(* IEC 61131-3 sources: Test-Git_ESME26/TestProgettoESME_26.fbsproj/PacDriveLib Migration/Motion/MultiCam/PDL_FB_MultiCam.fb.st^/Init, 2 files *)

(* ---- Init.meth.st ---- *)
METHOD PRIVATE Init : BOOL
VAR_INPUT
END_VAR

Init := FALSE;

//check axis
IF i_ifDrive = 0 THEN
	SetDiagOutput(	i_etDiag	:= GD.ET_Diag.InputParameterInvalid,
					i_etDiagExt := PDL_ET_DiagExt.DriveInvalid,
					i_sMsg		:= 'i_ifDrive - Invalid Interface');
	RETURN;

ELSIF iq_lencMaster = 0 THEN
	SetDiagOutput(	i_etDiag	:= GD.ET_Diag.InputParameterInvalid,
					i_etDiagExt := PDL_ET_DiagExt.DriveInvalid,
					i_sMsg		:= 'iq_lencMaster - Invalid Interface');
	RETURN;
ELSE
	//get IF_DriveConfig
	xSuccess := __QUERYINTERFACE(i_ifDrive, ifGetParentDevice);
	IF xSuccess AND ifGetParentDevice <> 0 THEN
		ifDeviceAccess := ifGetParentDevice.GetParentDevice();
		xSuccess := __QUERYINTERFACE( ifDeviceAccess, ifDriveConfigAccess );
		IF xSuccess AND ifDriveConfigAccess <> 0 THEN
			ifDriveConfig := ifDriveConfigAccess.DriveConfig;
		END_IF
	END_IF

	xSuccess := __QUERYINTERFACE(ifDeviceAccess, ifDeviceTreeObjectAccess);
	IF xSuccess THEN
		sDriveName := ifDeviceTreeObjectAccess.DeviceTreeObject.Name;
	ELSE
		sDriveName := 'Axis';
	END_IF

	fbHalt.Axis := i_ifDrive;
	fbStop.Axis := i_ifDrive;
	fbMoveAbsolute.Axis := i_ifDrive;
	fbCamIn.Slave := i_ifDrive;
	fbCamIn.Master := iq_lencMaster;
	fbCamIn2.Slave := i_ifDrive;
	fbCamIn2.Master := iq_lencMaster;

	xSlaveIsModulo := i_ifDrive.xIsModulo;

END_IF

//read cycle time
pstTaskInfo := __CURRENTTASK.pTaskInfo;
IF pstTaskInfo <> 0
THEN
	lrOwnPlcTaskInterval	:= DWORD_TO_LREAL(pstTaskInfo^.dwInterval) / 1000000.0; //usec to sec
	lrTSwitch				:= DINT_TO_LREAL(i_diTXend) / 1000.0 + lrOwnPlcTaskInterval;
ELSE
	SetDiagOutput(	i_etDiag	:= GD.ET_Diag.UnexpectedProgramBehavior,
					i_etDiagExt := PDL_ET_DiagExt.UnexpectedFeedback,
					i_sMsg		:= 'IecTaskGetInfo3 - reading cycle time failed');
	RETURN;
END_IF

Init := TRUE;

(* ---- RegisterLoggerPoint.meth.st ---- *)
METHOD PUBLIC RegisterLoggerPoint
VAR_INPUT
	i_ifParent		: APL.IF_LoggerPoint;
	i_sName			: STRING[80];
END_VAR
VAR_OUTPUT
	q_etDiag		: GD.ET_Diag := GD.ET_Diag.Ok;
	q_etDiagExt		: PDL_ET_DiagExt := PDL_ET_DiagExt.Ok;
END_VAR
VAR
	etDiagBuffer		: GD.ET_Diag;
	etDiagExtBufferAPL	: APL.ET_DiagExt;
END_VAR

THIS^.fbLoggerPoint.RegisterLoggerPoint(	i_ifParent		:= i_ifParent,
											i_sName			:= i_sName,
											i_sType			:= 'FB_MultiCam',
											i_sSource		:= 'PDL',
											q_etDiag		=> etDiagBuffer,
											q_etDiagExt		=> etDiagExtBufferAPL);

IF (etDiagBuffer <> GD.ET_Diag.Ok) THEN
	CASE etDiagExtBufferAPL OF
		APL.ET_DiagExt.ParentInvalid:
			q_etDiag := GD.ET_Diag.InputParameterInvalid;
			q_etDiagExt := PDL_ET_DiagExt.ParentInvalid;

		APL.ET_DiagExt.ParentNotRegistered:
			q_etDiag := GD.ET_Diag.InputParameterInvalid;
			q_etDiagExt := PDL_ET_DiagExt.ParentNotRegistered;

		APL.ET_DiagExt.MaxNumberOfLoggerPointsExeeded:
			q_etDiag := GD.ET_Diag.InputParameterInvalid;
			q_etDiagExt := PDL_ET_DiagExt.MaxNumberOfLoggerPointsExeeded;

	ELSE
		q_etDiag := GD.ET_Diag.UnexpectedProgramBehavior;
		q_etdiagExt := PDL_ET_DiagExt.UnexpectedDiagExt;
	END_CASE
END_IF
